(* IEC 61131-3 sources: volt/packages/volt-lsp-iec/test-corpus/awa-palletizer/Device/Plc Logic/Application/Library Manager/CAA FB Factory, 7 files *)

(* ---- ERROR.dut ---- *)
TYPE ERROR :
(
	NO_ERROR := 0,
	FIRST_ERROR := 1500,
	INVALID_PARAMETER := 1502,
	WRONG_INTERFACE := 1503,
	WRONG_INSTANCE_DATA := 1504,
	WRONG_POOL_SIZE := 1505,
	WRONG_INSTANCE_COUNT := 1506,
	NO_MEMORY := 1507,
	FIRST_MF := 1525,
	LAST_ERROR := 1549
);
END_TYPE

(* ---- IDATA.itf ---- *)
INTERFACE IDATA
END_INTERFACE

METHOD PRVCHECKDATAINST : BOOL
VAR_OUTPUT
	PDATA : POINTER TO InstanceData;
END_VAR
END_METHOD

(* ---- IFACTORY.itf ---- *)
INTERFACE IFACTORY
END_INTERFACE

METHOD PRVALLOCINSTMEM : CAA.HANDLE
VAR_OUTPUT
	EERROR : ERROR;
END_VAR
END_METHOD

METHOD PRVFREEINSTMEM : BOOL
VAR_INPUT
	HINST : CAA.HANDLE;
END_VAR
END_METHOD

METHOD PRVGETINSTPOINTER : CAA.PVOID
VAR_INPUT
	HINST : CAA.HANDLE;
END_VAR
END_METHOD

METHOD PRVINSERTINST : BOOL
VAR_INPUT
	ITFINST : IInstance;
END_VAR
END_METHOD

METHOD PRVINSTINIT : BOOL
VAR_INPUT
	ITFINST : IInstance;
	HINST : CAA.HANDLE;
	ITFDATA : IData;
END_VAR
VAR_OUTPUT
	EERROR : ERROR;
END_VAR
END_METHOD

METHOD PRVREMOVEINST : BOOL
VAR_INPUT
	ITFINST : IInstance;
END_VAR
END_METHOD

(* ---- IINSTANCE.itf ---- *)
INTERFACE IINSTANCE
END_INTERFACE

METHOD DISPOSE : BOOL
END_METHOD

METHOD PRVINSTINIT : ERROR
VAR_INPUT
	ITFDATA : IData;
END_VAR
END_METHOD

METHOD PRVINSTRELEASE : BOOL
END_METHOD

METHOD PRVINSTRETAIN : BOOL
END_METHOD

(* ---- FACTORYBASE.pou ---- *)
FUNCTION_BLOCK FACTORYBASE
VAR
	_HPOOL : CAA.HANDLE;
	_ITFINSTLIST : IInstance;
	_HPOOLSYNC : RTS_IEC_HANDLE := RTS_INVALID_HANDLE;
	_HLISTSYNC : RTS_IEC_HANDLE := RTS_INVALID_HANDLE;
	PRVINSTCOUNT : CAA.COUNT;
	PRVINSTPOOLADR : CAA.PVOID;
	PRVINSTPOOLEXTENDSFACTOR : USINT;
	PRVINSTPOOLSIZE : CAA.SIZE;
	PRVINSTSIZE : CAA.SIZE;
END_VAR
END_FUNCTION_BLOCK

METHOD FB_EXIT : BOOL
VAR_INPUT
	BINCOPYCODE : BOOL;
END_VAR
END_METHOD

METHOD FB_INIT : BOOL
VAR_INPUT
	BINITRETAINS : BOOL;
	BINCOPYCODE : BOOL;
END_VAR
END_METHOD

METHOD PRVALLOCINSTMEM : CAA.HANDLE
VAR_OUTPUT
	EERROR : ERROR;
END_VAR
END_METHOD

METHOD PRVFREEINSTMEM : BOOL
VAR_INPUT
	HINST : CAA.HANDLE;
END_VAR
END_METHOD

METHOD PRVGETINSTPOINTER : CAA.PVOID
VAR_INPUT
	HINST : CAA.HANDLE;
END_VAR
END_METHOD

METHOD PRVINSERTINST : BOOL
VAR_INPUT
	ITFINST : IInstance;
END_VAR
END_METHOD

METHOD PRVINSTINIT : BOOL
VAR_INPUT
	ITFINST : IInstance;
	HINST : CAA.HANDLE;
	ITFDATA : IData;
END_VAR
VAR_OUTPUT
	EERROR : ERROR;
END_VAR
END_METHOD

METHOD PRVREMOVEINST : BOOL
VAR_INPUT
	ITFINST : IInstance;
END_VAR
END_METHOD

(* ---- INSTANCEBASE.pou ---- *)
FUNCTION_BLOCK INSTANCEBASE
VAR
	_HINST : CAA.HANDLE;
	_ITFFACTORY : IFactory;
	_ITFNEXTINST : IInstance;
	_ITFPREVINST : IInstance;
	_CTREFCOUNT : CAA.COUNT;
	PRVINSTFACTORY : IFactory;
	PRVNEXTINST : IInstance;
	PRVPREVINST : IInstance;
END_VAR
END_FUNCTION_BLOCK

METHOD DISPOSE : BOOL
END_METHOD

METHOD PRVINSTINIT : ERROR
VAR_INPUT
	ITFDATA : IData;
END_VAR
END_METHOD

METHOD PRVINSTRELEASE : BOOL
END_METHOD

METHOD PRVINSTRETAIN : BOOL
END_METHOD

(* ---- INSTANCEDATA.pou ---- *)
FUNCTION_BLOCK INSTANCEDATA
VAR_INPUT
	HINST : CAA.HANDLE;
END_VAR
VAR
	C_DWDATASIGNATURE : DWORD := 16#68617461;
END_VAR
END_FUNCTION_BLOCK

METHOD PRVCHECKDATAINST : BOOL
VAR_OUTPUT
	PDATA : POINTER TO InstanceData;
END_VAR
END_METHOD
